(* IEC 61131-3 sources: plcfuzz/testcases/beremiz_projects/random_projects, 27 files *)

(* ---- G4LTL_ST1.st ---- *)
FUNCTION_BLOCK FB_G4LTL

   (* Variable definition *)
   VAR_INPUT
      x0	: BOOL;
      x1	: BOOL;
   END_VAR
   VAR_OUTPUT
      y0	: BOOL;
   END_VAR
   VAR
   (* The total number of states equals to 1 *)
      cstate0	: LINT := 0;
   END_VAR

   (* Control logic *)
CASE cstate0 OF
0:
    IF ((x0 = FALSE) AND  ( TRUE )) OR ((x0 = TRUE) AND  (x1 = TRUE)) THEN
        cstate0 := 0; y0 := FALSE;
    ELSIF ((x0 = TRUE) AND  (x1 = FALSE)) THEN
        cstate0 := 0; y0 := TRUE;
    END_IF;
END_CASE;

END_FUNCTION_BLOCK

(* ---- G4LTL_ST10.st ---- *)
FUNCTION_BLOCK FB_G4LTL

   (* Variable definition *)
   VAR_INPUT
      x1	: BOOL;
      x2	: BOOL;
   END_VAR
   VAR_OUTPUT
      y0	: BOOL;
      y1	: BOOL;
      y2	: BOOL;
   END_VAR
   VAR
   (* The total number of states equals to 6 *)
      cstate79	: LINT := 0;
   END_VAR

   (* Control logic *)
CASE cstate79 OF
0:
    IF ((x1 = FALSE) AND  (x2 = TRUE)) THEN
        cstate79 := 1; y0 := FALSE; y1 := FALSE; y2 := TRUE;
    ELSIF ((x1 = FALSE) AND  (x2 = FALSE)) THEN
        cstate79 := 2; y0 := FALSE; y1 := FALSE; y2 := TRUE;
    ELSIF ((x1 = TRUE) AND  (x2 = FALSE)) THEN
        cstate79 := 3; y0 := TRUE; y1 := TRUE; y2 := FALSE;
    ELSIF ((x1 = TRUE) AND  (x2 = TRUE)) THEN
        cstate79 := 5; y0 := FALSE; y1 := FALSE; y2 := FALSE;
    END_IF;
1:
    IF ((x1 = TRUE) AND  (x2 = FALSE)) THEN
        cstate79 := 3; y0 := TRUE; y1 := TRUE; y2 := FALSE;
    ELSIF ((x1 = TRUE) AND  (x2 = TRUE)) THEN
        cstate79 := 5; y0 := FALSE; y1 := FALSE; y2 := FALSE;
    ELSIF ((x1 = FALSE) AND  ( TRUE )) THEN
        cstate79 := 1; y0 := FALSE; y1 := FALSE; y2 := TRUE;
    END_IF;
2:
    IF ((x1 = TRUE) AND  (x2 = FALSE)) THEN
        cstate79 := 3; y0 := TRUE; y1 := TRUE; y2 := FALSE;
    ELSIF ((x1 = FALSE) AND  (x2 = TRUE)) THEN
        cstate79 := 1; y0 := FALSE; y1 := FALSE; y2 := TRUE;
    ELSIF ((x1 = TRUE) AND  (x2 = TRUE)) THEN
        cstate79 := 5; y0 := FALSE; y1 := FALSE; y2 := FALSE;
    ELSIF ((x1 = FALSE) AND  (x2 = FALSE)) THEN
        cstate79 := 2; y0 := FALSE; y1 := FALSE; y2 := TRUE;
    END_IF;
3:
    IF ((x1 = FALSE) AND  (x2 = TRUE)) THEN
        cstate79 := 4; y0 := FALSE; y1 := FALSE; y2 := TRUE;
    ELSIF (( TRUE ) AND  (x2 = FALSE)) THEN
        cstate79 := 3; y0 := TRUE; y1 := TRUE; y2 := FALSE;
    ELSIF ((x1 = TRUE) AND  (x2 = TRUE)) THEN
        cstate79 := 5; y0 := FALSE; y1 := FALSE; y2 := FALSE;
    END_IF;
4:
    IF ((x1 = TRUE) AND  (x2 = FALSE)) THEN
        cstate79 := 3; y0 := TRUE; y1 := TRUE; y2 := FALSE;
    ELSIF ((x1 = TRUE) AND  (x2 = TRUE)) THEN
        cstate79 := 5; y0 := FALSE; y1 := FALSE; y2 := FALSE;
    ELSIF ((x1 = FALSE) AND  ( TRUE )) THEN
        cstate79 := 4; y0 := FALSE; y1 := FALSE; y2 := TRUE;
    END_IF;
5:
    IF ((x1 = FALSE) AND  (x2 = FALSE)) THEN
        cstate79 := 5; y0 := FALSE; y1 := FALSE; y2 := FALSE;
    ELSIF ((x1 = TRUE) AND  (x2 = TRUE)) THEN
        cstate79 := 5; y0 := FALSE; y1 := FALSE; y2 := FALSE;
    ELSIF ((x1 = TRUE) AND  (x2 = FALSE)) THEN
        cstate79 := 3; y0 := TRUE; y1 := TRUE; y2 := FALSE;
    ELSIF ((x1 = FALSE) AND  (x2 = TRUE)) THEN
        cstate79 := 4; y0 := FALSE; y1 := FALSE; y2 := TRUE;
    END_IF;
END_CASE;

END_FUNCTION_BLOCK

(* ---- G4LTL_ST2.st ---- *)
FUNCTION_BLOCK FB_G4LTL

   (* Variable definition *)
   VAR_INPUT
      x0	: BOOL;
      x1	: BOOL;
   END_VAR
   VAR_OUTPUT
      y0	: BOOL;
   END_VAR
   VAR
   (* The total number of states equals to 1 *)
      cstate99	: LINT := 0;
   END_VAR

   (* Control logic *)
CASE cstate99 OF
0:
    IF ((x0 = FALSE) AND  (x1 = TRUE)) OR ((x0 = TRUE) AND  (x1 = FALSE)) THEN
        cstate99 := 0; y0 := FALSE;
    ELSIF ((x0 = FALSE) AND  (x1 = FALSE)) OR ((x0 = TRUE) AND  (x1 = TRUE)) THEN
        cstate99 := 0; y0 := TRUE;
    END_IF;
END_CASE;

END_FUNCTION_BLOCK

(* ---- G4LTL_ST3.st ---- *)
FUNCTION_BLOCK FB_G4LTL

   (* Variable definition *)
   VAR_INPUT
      x0	: BOOL;
      x1	: BOOL;
      x2	: BOOL;
      x3	: BOOL;
   END_VAR
   VAR_OUTPUT
      y0	: BOOL;
   END_VAR
   VAR
   (* The total number of states equals to 12 *)
      cstate33	: LINT := 0;
   END_VAR

   (* Control logic *)
CASE cstate33 OF
22:
    IF ((x0 = TRUE) AND  (x1 = TRUE) AND  (x2 = TRUE) AND  (x3 = FALSE)) THEN
        cstate33 := 247; y0 := FALSE;
    ELSIF ((x0 = FALSE) AND  ( TRUE ) AND  ( TRUE ) AND  ( TRUE )) OR ((x0 = TRUE) AND  ( TRUE ) AND  (x2 = FALSE) AND  ( TRUE )) THEN
        cstate33 := 22; y0 := FALSE;
    ELSIF ((x0 = TRUE) AND  (x1 = FALSE) AND  (x2 = TRUE) AND  (x3 = FALSE)) THEN
        cstate33 := 246; y0 := TRUE;
    ELSIF ((x0 = TRUE) AND  ( TRUE ) AND  (x2 = TRUE) AND  (x3 = TRUE)) THEN
        cstate33 := 29; y0 := FALSE;
    END_IF;
0:
    IF ((x0 = FALSE) AND  (x1 = FALSE) AND  (x2 = TRUE) AND  (x3 = FALSE)) THEN
        cstate33 := 0; y0 := FALSE;
    ELSIF ((x0 = FALSE) AND  (x1 = TRUE) AND  (x2 = TRUE) AND  (x3 = FALSE)) THEN
        cstate33 := 24; y0 := FALSE;
    ELSIF ((x0 = FALSE) AND  (x1 = TRUE) AND  ( TRUE ) AND  (x3 = TRUE)) OR ((x0 = TRUE) AND  (x1 = TRUE) AND  (x2 = FALSE) AND  (x3 = TRUE)) THEN
        cstate33 := 22; y0 := FALSE;
    ELSIF ((x0 = TRUE) AND  (x1 = TRUE) AND  (x2 = TRUE) AND  (x3 = FALSE)) THEN
        cstate33 := 28; y0 := FALSE;
    ELSIF (( TRUE ) AND  (x1 = TRUE) AND  (x2 = FALSE) AND  (x3 = FALSE)) THEN
        cstate33 := 20; y0 := FALSE;
    ELSIF ((x0 = TRUE) AND  (x1 = FALSE) AND  (x2 = TRUE) AND  (x3 = FALSE)) THEN
        cstate33 := 27; y0 := TRUE;
    ELSIF ((x0 = TRUE) AND  (x1 = TRUE) AND  (x2 = TRUE) AND  (x3 = TRUE)) THEN
        cstate33 := 29; y0 := FALSE;
    ELSIF (( TRUE ) AND  (x1 = FALSE) AND  (x2 = FALSE) AND  ( TRUE )) OR (( TRUE ) AND  (x1 = FALSE) AND  (x2 = TRUE) AND  (x3 = TRUE)) THEN
        cstate33 := 18; y0 := FALSE;
    END_IF;
243:
    IF ((x0 = FALSE) AND  (x1 = FALSE) AND  (x2 = TRUE) AND  (x3 = TRUE)) OR ((x0 = TRUE) AND  ( TRUE ) AND  (x2 = TRUE) AND  (x3 = TRUE)) THEN
        cstate33 := 29; y0 := FALSE;
    ELSIF (( TRUE ) AND  ( TRUE ) AND  (x2 = FALSE) AND  (x3 = FALSE)) THEN
        cstate33 := 20; y0 := FALSE;
    ELSIF ((x0 = FALSE) AND  (x1 = FALSE) AND  (x2 = FALSE) AND  (x3 = TRUE)) OR ((x0 = FALSE) AND  (x1 = TRUE) AND  ( TRUE ) AND  (x3 = TRUE)) OR ((x0 = TRUE) AND  ( TRUE ) AND  (x2 = FALSE) AND  (x3 = TRUE)) THEN
        cstate33 := 22; y0 := FALSE;
    ELSIF ((x0 = FALSE) AND  (x1 = TRUE) AND  (x2 = TRUE) AND  (x3 = FALSE)) THEN
        cstate33 := 24; y0 := FALSE;
    ELSIF ((x0 = TRUE) AND  (x1 = TRUE) AND  (x2 = TRUE) AND  (x3 = FALSE)) THEN
        cstate33 := 28; y0 := FALSE;
    ELSIF (( TRUE ) AND  (x1 = FALSE) AND  (x2 = TRUE) AND  (x3 = FALSE)) THEN
        cstate33 := 243; y0 := TRUE;
    END_IF;
24:
    IF ((x0 = TRUE) AND  ( TRUE ) AND  (x2 = TRUE) AND  (x3 = TRUE)) THEN
        cstate33 := 29; y0 := FALSE;
    ELSIF (( TRUE ) AND  ( TRUE ) AND  (x2 = FALSE) AND  (x3 = FALSE)) THEN
        cstate33 := 20; y0 := FALSE;
    ELSIF ((x0 = FALSE) AND  ( TRUE ) AND  ( TRUE ) AND  (x3 = TRUE)) OR ((x0 = TRUE) AND  ( TRUE ) AND  (x2 = FALSE) AND  (x3 = TRUE)) THEN
        cstate33 := 22; y0 := FALSE;
    ELSIF ((x0 = TRUE) AND  (x1 = TRUE) AND  (x2 = TRUE) AND  (x3 = FALSE)) THEN
        cstate33 := 28; y0 := FALSE;
    ELSIF ((x0 = TRUE) AND  (x1 = FALSE) AND  (x2 = TRUE) AND  (x3 = FALSE)) THEN
        cstate33 := 243; y0 := TRUE;
    ELSIF ((x0 = FALSE) AND  ( TRUE ) AND  (x2 = TRUE) AND  (x3 = FALSE)) THEN
        cstate33 := 24; y0 := FALSE;
    END_IF;
246:
    IF ((x0 = FALSE) AND  (x1 = FALSE) AND  (x2 = FALSE) AND  ( TRUE )) OR ((x0 = FALSE) AND  (x1 = TRUE) AND  (x2 = FALSE) AND  ( TRUE )) OR ((x0 = FALSE) AND  (x1 = TRUE) AND  (x2 = TRUE) AND  (x3 = TRUE)) OR ((x0 = TRUE) AND  ( TRUE ) AND  (x2 = FALSE) AND  ( TRUE )) THEN
        cstate33 := 22; y0 := FALSE;
    ELSIF (( TRUE ) AND  (x1 = FALSE) AND  (x2 = TRUE) AND  (x3 = FALSE)) THEN
        cstate33 := 246; y0 := TRUE;
    ELSIF ((x0 = FALSE) AND  (x1 = FALSE) AND  (x2 = TRUE) AND  (x3 = TRUE)) OR ((x0 = TRUE) AND  ( TRUE ) AND  (x2 = TRUE) AND  (x3 = TRUE)) THEN
        cstate33 := 29; y0 := FALSE;
    ELSIF ((x0 = FALSE) AND  (x1 = TRUE) AND  (x2 = TRUE) AND  (x3 = FALSE)) THEN
        cstate33 := 786; y0 := FALSE;
    ELSIF ((x0 = TRUE) AND  (x1 = TRUE) AND  (x2 = TRUE) AND  (x3 = FALSE)) THEN
        cstate33 := 247; y0 := FALSE;
    END_IF;
27:
    IF ((x0 = FALSE) AND  (x1 = TRUE) AND  (x2 = TRUE) AND  (x3 = FALSE)) THEN
        cstate33 := 24; y0 := FALSE;
    ELSIF (( TRUE ) AND  (x1 = TRUE) AND  (x2 = FALSE) AND  (x3 = FALSE)) THEN
        cstate33 := 20; y0 := FALSE;
    ELSIF ((x0 = FALSE) AND  (x1 = TRUE) AND  ( TRUE ) AND  (x3 = TRUE)) OR ((x0 = TRUE) AND  (x1 = TRUE) AND  (x2 = FALSE) AND  (x3 = TRUE)) THEN
        cstate33 := 22; y0 := FALSE;
    ELSIF ((x0 = TRUE) AND  (x1 = TRUE) AND  (x2 = TRUE) AND  (x3 = FALSE)) THEN
        cstate33 := 28; y0 := FALSE;
    ELSIF (( TRUE ) AND  (x1 = FALSE) AND  (x2 = TRUE) AND  (x3 = FALSE)) THEN
        cstate33 := 27; y0 := TRUE;
    ELSIF ((x0 = TRUE) AND  (x1 = TRUE) AND  (x2 = TRUE) AND  (x3 = TRUE)) THEN
        cstate33 := 29; y0 := FALSE;
    ELSIF (( TRUE ) AND  (x1 = FALSE) AND  (x2 = FALSE) AND  ( TRUE )) OR (( TRUE ) AND  (x1 = FALSE) AND  (x2 = TRUE) AND  (x3 = TRUE)) THEN
        cstate33 := 18; y0 := FALSE;
    END_IF;
247:
    IF ((x0 = FALSE) AND  (x1 = TRUE) AND  (x2 = TRUE) AND  (x3 = FALSE)) THEN
        cstate33 := 786; y0 := FALSE;
    ELSIF ((x0 = FALSE) AND  (x1 = FALSE) AND  (x2 = TRUE) AND  (x3 = FALSE)) OR ((x0 = TRUE) AND  (x1 = TRUE) AND  (x2 = TRUE) AND  (x3 = FALSE)) THEN
        cstate33 := 247; y0 := FALSE;
    ELSIF ((x0 = FALSE) AND  (x1 = FALSE) AND  (x2 = FALSE) AND  ( TRUE )) OR ((x0 = FALSE) AND  (x1 = TRUE) AND  (x2 = FALSE) AND  ( TRUE )) OR ((x0 = FALSE) AND  (x1 = TRUE) AND  (x2 = TRUE) AND  (x3 = TRUE)) OR ((x0 = TRUE) AND  ( TRUE ) AND  (x2 = FALSE) AND  ( TRUE )) THEN
        cstate33 := 22; y0 := FALSE;
    ELSIF ((x0 = TRUE) AND  (x1 = FALSE) AND  (x2 = TRUE) AND  (x3 = FALSE)) THEN
        cstate33 := 246; y0 := TRUE;
    ELSIF ((x0 = FALSE) AND  (x1 = FALSE) AND  (x2 = TRUE) AND  (x3 = TRUE)) OR ((x0 = TRUE) AND  ( TRUE ) AND  (x2 = TRUE) AND  (x3 = TRUE)) THEN
        cstate33 := 29; y0 := FALSE;
    END_IF;
786:
    IF ((x0 = TRUE) AND  (x1 = TRUE) AND  (x2 = TRUE) AND  (x3 = FALSE)) THEN
        cstate33 := 247; y0 := FALSE;
    ELSIF ((x0 = FALSE) AND  ( TRUE ) AND  (x2 = FALSE) AND  ( TRUE )) OR ((x0 = FALSE) AND  ( TRUE ) AND  (x2 = TRUE) AND  (x3 = TRUE)) OR ((x0 = TRUE) AND  ( TRUE ) AND  (x2 = FALSE) AND  ( TRUE )) THEN
        cstate33 := 22; y0 := FALSE;
    ELSIF ((x0 = FALSE) AND  ( TRUE ) AND  (x2 = TRUE) AND  (x3 = FALSE)) THEN
        cstate33 := 786; y0 := FALSE;
    ELSIF ((x0 = TRUE) AND  (x1 = FALSE) AND  (x2 = TRUE) AND  (x3 = FALSE)) THEN
        cstate33 := 246; y0 := TRUE;
    ELSIF ((x0 = TRUE) AND  ( TRUE ) AND  (x2 = TRUE) AND  (x3 = TRUE)) THEN
        cstate33 := 29; y0 := FALSE;
    END_IF;
28:
    IF ((x0 = FALSE) AND  (x1 = FALSE) AND  (x2 = TRUE) AND  (x3 = FALSE)) OR ((x0 = TRUE) AND  (x1 = TRUE) AND  (x2 = TRUE) AND  (x3 = FALSE)) THEN
        cstate33 := 28; y0 := FALSE;
    ELSIF (( TRUE ) AND  ( TRUE ) AND  (x2 = FALSE) AND  (x3 = FALSE)) THEN
        cstate33 := 20; y0 := FALSE;
    ELSIF ((x0 = FALSE) AND  (x1 = FALSE) AND  (x2 = FALSE) AND  (x3 = TRUE)) OR ((x0 = FALSE) AND  (x1 = TRUE) AND  ( TRUE ) AND  (x3 = TRUE)) OR ((x0 = TRUE) AND  ( TRUE ) AND  (x2 = FALSE) AND  (x3 = TRUE)) THEN
        cstate33 := 22; y0 := FALSE;
    ELSIF ((x0 = FALSE) AND  (x1 = TRUE) AND  (x2 = TRUE) AND  (x3 = FALSE)) THEN
        cstate33 := 24; y0 := FALSE;
    ELSIF ((x0 = TRUE) AND  (x1 = FALSE) AND  (x2 = TRUE) AND  (x3 = FALSE)) THEN
        cstate33 := 243; y0 := TRUE;
    ELSIF ((x0 = FALSE) AND  (x1 = FALSE) AND  (x2 = TRUE) AND  (x3 = TRUE)) OR ((x0 = TRUE) AND  ( TRUE ) AND  (x2 = TRUE) AND  (x3 = TRUE)) THEN
        cstate33 := 29; y0 := FALSE;
    END_IF;
29:
    IF ((x0 = TRUE) AND  (x1 = TRUE) AND  (x2 = TRUE) AND  (x3 = FALSE)) THEN
        cstate33 := 247; y0 := FALSE;
    ELSIF ((x0 = FALSE) AND  (x1 = FALSE) AND  (x2 = TRUE) AND  ( TRUE )) OR ((x0 = TRUE) AND  ( TRUE ) AND  (x2 = TRUE) AND  (x3 = TRUE)) THEN
        cstate33 := 29; y0 := FALSE;
    ELSIF ((x0 = TRUE) AND  (x1 = FALSE) AND  (x2 = TRUE) AND  (x3 = FALSE)) THEN
        cstate33 := 246; y0 := TRUE;
    ELSIF ((x0 = FALSE) AND  (x1 = FALSE) AND  (x2 = FALSE) AND  ( TRUE )) OR ((x0 = FALSE) AND  (x1 = TRUE) AND  ( TRUE ) AND  ( TRUE )) OR ((x0 = TRUE) AND  ( TRUE ) AND  (x2 = FALSE) AND  ( TRUE )) THEN
        cstate33 := 22; y0 := FALSE;
    END_IF;
18:
    IF ((x0 = TRUE) AND  (x1 = TRUE) AND  (x2 = TRUE) AND  (x3 = TRUE)) THEN
        cstate33 := 29; y0 := FALSE;
    ELSIF ((x0 = TRUE) AND  (x1 = FALSE) AND  (x2 = TRUE) AND  (x3 = FALSE)) THEN
        cstate33 := 27; y0 := TRUE;
    ELSIF ((x0 = FALSE) AND  (x1 = FALSE) AND  ( TRUE ) AND  ( TRUE )) OR ((x0 = TRUE) AND  (x1 = FALSE) AND  (x2 = FALSE) AND  ( TRUE )) OR ((x0 = TRUE) AND  (x1 = FALSE) AND  (x2 = TRUE) AND  (x3 = TRUE)) THEN
        cstate33 := 18; y0 := FALSE;
    ELSIF ((x0 = FALSE) AND  (x1 = TRUE) AND  ( TRUE ) AND  (x3 = FALSE)) OR ((x0 = TRUE) AND  (x1 = TRUE) AND  (x2 = FALSE) AND  (x3 = FALSE)) THEN
        cstate33 := 20; y0 := FALSE;
    ELSIF ((x0 = FALSE) AND  (x1 = TRUE) AND  ( TRUE ) AND  (x3 = TRUE)) OR ((x0 = TRUE) AND  (x1 = TRUE) AND  (x2 = FALSE) AND  (x3 = TRUE)) THEN
        cstate33 := 22; y0 := FALSE;
    ELSIF ((x0 = TRUE) AND  (x1 = TRUE) AND  (x2 = TRUE) AND  (x3 = FALSE)) THEN
        cstate33 := 28; y0 := FALSE;
    END_IF;
20:
    IF ((x0 = TRUE) AND  ( TRUE ) AND  (x2 = TRUE) AND  (x3 = TRUE)) THEN
        cstate33 := 29; y0 := FALSE;
    ELSIF ((x0 = FALSE) AND  ( TRUE ) AND  ( TRUE ) AND  (x3 = TRUE)) OR ((x0 = TRUE) AND  ( TRUE ) AND  (x2 = FALSE) AND  (x3 = TRUE)) THEN
        cstate33 := 22; y0 := FALSE;
    ELSIF ((x0 = FALSE) AND  ( TRUE ) AND  ( TRUE ) AND  (x3 = FALSE)) OR ((x0 = TRUE) AND  ( TRUE ) AND  (x2 = FALSE) AND  (x3 = FALSE)) THEN
        cstate33 := 20; y0 := FALSE;
    ELSIF ((x0 = TRUE) AND  (x1 = TRUE) AND  (x2 = TRUE) AND  (x3 = FALSE)) THEN
        cstate33 := 28; y0 := FALSE;
    ELSIF ((x0 = TRUE) AND  (x1 = FALSE) AND  (x2 = TRUE) AND  (x3 = FALSE)) THEN
        cstate33 := 243; y0 := TRUE;
    END_IF;
END_CASE;

END_FUNCTION_BLOCK

(* ---- G4LTL_ST4.st ---- *)
FUNCTION_BLOCK FB_G4LTL

   (* Variable definition *)
   VAR_INPUT
      x0	: BOOL;
      x1	: BOOL;
      x2	: BOOL;
      x3	: BOOL;
   END_VAR
   VAR_OUTPUT
      y0	: BOOL;
      y1	: BOOL;
   END_VAR
   VAR
   (* The total number of states equals to 2 *)
      cstate29	: LINT := 0;
   END_VAR

   (* Control logic *)
CASE cstate29 OF
0:
    IF ((x0 = FALSE) AND  (x1 = FALSE) AND  (x2 = FALSE) AND  (x3 = TRUE)) THEN
        cstate29 := 0; y0 := FALSE; y1 := FALSE;
    ELSIF ((x0 = FALSE) AND  (x1 = TRUE) AND  ( TRUE ) AND  (x3 = TRUE)) OR ((x0 = TRUE) AND  (x1 = FALSE) AND  (x2 = TRUE) AND  ( TRUE )) OR ((x0 = TRUE) AND  (x1 = TRUE) AND  (x2 = FALSE) AND  (x3 = TRUE)) OR ((x0 = TRUE) AND  (x1 = TRUE) AND  (x2 = TRUE) AND  ( TRUE )) THEN
        cstate29 := 1; y0 := FALSE; y1 := FALSE;
    ELSIF ((x0 = FALSE) AND  (x1 = FALSE) AND  (x2 = FALSE) AND  (x3 = FALSE)) OR ((x0 = FALSE) AND  (x1 = FALSE) AND  (x2 = TRUE) AND  ( TRUE )) OR ((x0 = FALSE) AND  (x1 = TRUE) AND  ( TRUE ) AND  (x3 = FALSE)) THEN
        cstate29 := 0; y0 := FALSE; y1 := FALSE;
    ELSIF ((x0 = TRUE) AND  (x1 = TRUE) AND  (x2 = FALSE) AND  (x3 = FALSE)) THEN
        cstate29 := 0; y0 := TRUE; y1 := TRUE;
    ELSIF ((x0 = TRUE) AND  (x1 = FALSE) AND  (x2 = FALSE) AND  (x3 = TRUE)) THEN
        cstate29 := 0; y0 := TRUE; y1 := FALSE;
    ELSIF ((x0 = TRUE) AND  (x1 = FALSE) AND  (x2 = FALSE) AND  (x3 = FALSE)) THEN
        cstate29 := 0; y0 := TRUE; y1 := FALSE;
    END_IF;
1:
    IF ((x0 = TRUE) AND  (x1 = FALSE) AND  (x2 = FALSE) AND  ( TRUE )) OR ((x0 = TRUE) AND  (x1 = TRUE) AND  (x2 = FALSE) AND  (x3 = FALSE)) THEN
        cstate29 := 1; y0 := FALSE; y1 := FALSE;
    ELSIF ((x0 = FALSE) AND  (x1 = FALSE) AND  (x2 = FALSE) AND  (x3 = FALSE)) OR ((x0 = FALSE) AND  (x1 = FALSE) AND  (x2 = TRUE) AND  ( TRUE )) OR ((x0 = FALSE) AND  (x1 = TRUE) AND  ( TRUE ) AND  (x3 = FALSE)) THEN
        cstate29 := 1; y0 := FALSE; y1 := FALSE;
    ELSIF ((x0 = FALSE) AND  (x1 = TRUE) AND  ( TRUE ) AND  (x3 = TRUE)) OR ((x0 = TRUE) AND  (x1 = FALSE) AND  (x2 = TRUE) AND  ( TRUE )) OR ((x0 = TRUE) AND  (x1 = TRUE) AND  (x2 = FALSE) AND  (x3 = TRUE)) OR ((x0 = TRUE) AND  (x1 = TRUE) AND  (x2 = TRUE) AND  ( TRUE )) THEN
        cstate29 := 1; y0 := FALSE; y1 := FALSE;
    ELSIF ((x0 = FALSE) AND  (x1 = FALSE) AND  (x2 = FALSE) AND  (x3 = TRUE)) THEN
        cstate29 := 1; y0 := FALSE; y1 := FALSE;
    END_IF;
END_CASE;

END_FUNCTION_BLOCK

(* ---- G4LTL_ST5.st ---- *)
FUNCTION_BLOCK FB_G4LTL

   (* Variable definition *)
   VAR_INPUT
      x0	: BOOL;
      x1	: BOOL;
      c1_geq500	: BOOL;
   END_VAR
   VAR_OUTPUT
      y0	: BOOL;
      c1_add1	: BOOL;
      c1_reset	: BOOL;
   END_VAR
   VAR
   (* The total number of states equals to 4 *)
      cstate69	: LINT := 0;
   END_VAR

   (* Control logic *)
CASE cstate69 OF
0:
    IF ((x0 = FALSE) AND  (x1 = TRUE) AND  (c1_geq500 = TRUE)) THEN
        cstate69 := 3; y0 := TRUE; c1_add1 := FALSE; c1_reset := TRUE;
    ELSIF ((x0 = FALSE) AND  (x1 = FALSE) AND  (c1_geq500 = TRUE)) THEN
        cstate69 := 3; y0 := TRUE; c1_add1 := FALSE; c1_reset := FALSE;
    ELSIF ((x0 = FALSE) AND  (x1 = TRUE) AND  (c1_geq500 = FALSE)) THEN
        cstate69 := 3; y0 := FALSE; c1_add1 := FALSE; c1_reset := TRUE;
    ELSIF ((x0 = FALSE) AND  (x1 = FALSE) AND  (c1_geq500 = FALSE)) THEN
        cstate69 := 3; y0 := FALSE; c1_add1 := FALSE; c1_reset := FALSE;
    ELSIF ((x0 = TRUE) AND  (x1 = TRUE) AND  ( TRUE )) THEN
        cstate69 := 1; y0 := FALSE; c1_add1 := FALSE; c1_reset := FALSE;
    ELSIF ((x0 = TRUE) AND  (x1 = FALSE) AND  (c1_geq500 = TRUE)) THEN
        cstate69 := 2; y0 := TRUE; c1_add1 := TRUE; c1_reset := FALSE;
    ELSIF ((x0 = TRUE) AND  (x1 = FALSE) AND  (c1_geq500 = FALSE)) THEN
        cstate69 := 2; y0 := FALSE; c1_add1 := TRUE; c1_reset := FALSE;
    END_IF;
1:
    IF ((x0 = TRUE) AND  (x1 = TRUE) AND  ( TRUE )) THEN
        cstate69 := 1; y0 := FALSE; c1_add1 := FALSE; c1_reset := FALSE;
    ELSIF ((x0 = FALSE) AND  ( TRUE ) AND  (c1_geq500 = FALSE)) OR ((x0 = TRUE) AND  (x1 = FALSE) AND  (c1_geq500 = FALSE)) THEN
        cstate69 := 1; y0 := FALSE; c1_add1 := FALSE; c1_reset := FALSE;
    ELSIF ((x0 = FALSE) AND  ( TRUE ) AND  (c1_geq500 = TRUE)) OR ((x0 = TRUE) AND  (x1 = FALSE) AND  (c1_geq500 = TRUE)) THEN
        cstate69 := 1; y0 := FALSE; c1_add1 := FALSE; c1_reset := FALSE;
    END_IF;
2:
    IF ((x0 = TRUE) AND  (x1 = TRUE) AND  ( TRUE )) THEN
        cstate69 := 1; y0 := FALSE; c1_add1 := FALSE; c1_reset := FALSE;
    ELSIF ((x0 = FALSE) AND  (x1 = FALSE) AND  (c1_geq500 = TRUE)) THEN
        cstate69 := 3; y0 := TRUE; c1_add1 := FALSE; c1_reset := FALSE;
    ELSIF ((x0 = FALSE) AND  (x1 = TRUE) AND  (c1_geq500 = FALSE)) THEN
        cstate69 := 3; y0 := FALSE; c1_add1 := FALSE; c1_reset := TRUE;
    ELSIF ((x0 = FALSE) AND  (x1 = TRUE) AND  (c1_geq500 = TRUE)) THEN
        cstate69 := 3; y0 := TRUE; c1_add1 := FALSE; c1_reset := TRUE;
    ELSIF ((x0 = FALSE) AND  (x1 = FALSE) AND  (c1_geq500 = FALSE)) THEN
        cstate69 := 3; y0 := FALSE; c1_add1 := FALSE; c1_reset := FALSE;
    ELSIF ((x0 = TRUE) AND  (x1 = FALSE) AND  (c1_geq500 = FALSE)) THEN
        cstate69 := 2; y0 := FALSE; c1_add1 := FALSE; c1_reset := FALSE;
    ELSIF ((x0 = TRUE) AND  (x1 = FALSE) AND  (c1_geq500 = TRUE)) THEN
        cstate69 := 2; y0 := TRUE; c1_add1 := FALSE; c1_reset := FALSE;
    END_IF;
3:
    IF ((x0 = FALSE) AND  (x1 = FALSE) AND  (c1_geq500 = FALSE)) THEN
        cstate69 := 3; y0 := FALSE; c1_add1 := FALSE; c1_reset := FALSE;
    ELSIF ((x0 = FALSE) AND  (x1 = FALSE) AND  (c1_geq500 = TRUE)) THEN
        cstate69 := 3; y0 := TRUE; c1_add1 := FALSE; c1_reset := FALSE;
    ELSIF ((x0 = FALSE) AND  (x1 = TRUE) AND  (c1_geq500 = FALSE)) THEN
        cstate69 := 3; y0 := FALSE; c1_add1 := FALSE; c1_reset := TRUE;
    ELSIF ((x0 = FALSE) AND  (x1 = TRUE) AND  (c1_geq500 = TRUE)) THEN
        cstate69 := 3; y0 := TRUE; c1_add1 := FALSE; c1_reset := TRUE;
    ELSIF ((x0 = TRUE) AND  (x1 = TRUE) AND  ( TRUE )) THEN
        cstate69 := 1; y0 := FALSE; c1_add1 := FALSE; c1_reset := FALSE;
    ELSIF ((x0 = TRUE) AND  (x1 = FALSE) AND  (c1_geq500 = FALSE)) THEN
        cstate69 := 2; y0 := FALSE; c1_add1 := TRUE; c1_reset := FALSE;
    ELSIF ((x0 = TRUE) AND  (x1 = FALSE) AND  (c1_geq500 = TRUE)) THEN
        cstate69 := 2; y0 := TRUE; c1_add1 := TRUE; c1_reset := FALSE;
    END_IF;
END_CASE;

END_FUNCTION_BLOCK

(* ---- G4LTL_ST6.st ---- *)
FUNCTION_BLOCK FB_G4LTL

   (* Variable definition *)
   VAR_INPUT
      x1	: BOOL;
   END_VAR
   VAR_OUTPUT
      y1	: BOOL;
   END_VAR
   VAR
   (* The total number of states equals to 7 *)
      cstate14	: LINT := 0;
      t	: TON;
      t_reset	: BOOL := FALSE;
      t_up	: BOOL := FALSE;
      t_start	: BOOL := FALSE;
   END_VAR

   (* Constant definition (depending on compiler, one might need to move to normal variables) *)

   (* Each time constant has a difference of 1 period (cycle-time); please substract it when needed  *)
   VAR CONST
      T_VALUE	: TIME := TIME#5s;
   END_VAR

   (* Control logic *)
CASE cstate14 OF
0:
    IF ((x1 = FALSE) AND  (t.Q = FALSE)) THEN
        cstate14 := 1; y1 := FALSE; t_start := FALSE;
    ELSIF ((x1 = TRUE) AND  ( TRUE )) THEN
        cstate14 := 3; y1 := TRUE; t_start := FALSE;
    ELSIF ((x1 = FALSE) AND  (t.Q = TRUE)) THEN
        cstate14 := 5; y1 := FALSE; t_start := FALSE;
    END_IF;
1:
    IF ((x1 = FALSE) AND  (t.Q = FALSE)) THEN
        cstate14 := 1; y1 := FALSE; t_start := FALSE;
    ELSIF ((x1 = FALSE) AND  (t.Q = TRUE)) THEN
        cstate14 := 5; y1 := FALSE; t_start := FALSE;
    ELSIF ((x1 = TRUE) AND  ( TRUE )) THEN
        cstate14 := 3; y1 := TRUE; t_start := FALSE;
    END_IF;
2:
    IF ((x1 = TRUE) AND  (t.Q = FALSE)) THEN
        cstate14 := 2; y1 := TRUE; t_start := FALSE;
    ELSIF ((x1 = TRUE) AND  (t.Q = TRUE)) THEN
        cstate14 := 3; y1 := TRUE; t_start := FALSE;
    ELSIF ((x1 = FALSE) AND  (t.Q = FALSE)) THEN
        cstate14 := 4; y1 := TRUE; t_start := TRUE; t_up := FALSE;
    ELSIF ((x1 = FALSE) AND  (t.Q = TRUE)) THEN
        cstate14 := 6; y1 := TRUE; t_start := TRUE; t_up := FALSE;
    END_IF;
3:
    IF ((x1 = FALSE) AND  (t.Q = TRUE)) THEN
        cstate14 := 6; y1 := TRUE; t_start := TRUE; t_up := FALSE;
    ELSIF ((x1 = FALSE) AND  (t.Q = FALSE)) THEN
        cstate14 := 4; y1 := TRUE; t_start := TRUE; t_up := FALSE;
    ELSIF ((x1 = TRUE) AND  ( TRUE )) THEN
        cstate14 := 3; y1 := TRUE; t_start := FALSE;
    END_IF;
4:
    IF ((x1 = FALSE) AND  (t.Q = TRUE)) THEN
        cstate14 := 5; y1 := FALSE; t_start := FALSE;
    ELSIF ((x1 = FALSE) AND  (t.Q = FALSE)) THEN
        cstate14 := 4; y1 := TRUE; t_start := FALSE;
    ELSIF ((x1 = TRUE) AND  (t.Q = FALSE)) THEN
        cstate14 := 2; y1 := TRUE; t_start := FALSE;
    ELSIF ((x1 = TRUE) AND  (t.Q = TRUE)) THEN
        cstate14 := 3; y1 := TRUE; t_start := FALSE;
    END_IF;
5:
    IF ((x1 = TRUE) AND  ( TRUE )) THEN
        cstate14 := 3; y1 := TRUE; t_start := FALSE;
    ELSIF ((x1 = FALSE) AND  (t.Q = FALSE)) THEN
        cstate14 := 1; y1 := FALSE; t_start := FALSE;
    ELSIF ((x1 = FALSE) AND  (t.Q = TRUE)) THEN
        cstate14 := 5; y1 := FALSE; t_start := FALSE;
    END_IF;
6:
    IF ((x1 = FALSE) AND  (t.Q = TRUE)) THEN
        cstate14 := 5; y1 := FALSE; t_start := FALSE;
    ELSIF ((x1 = FALSE) AND  (t.Q = FALSE)) THEN
        cstate14 := 4; y1 := TRUE; t_start := FALSE;
    ELSIF ((x1 = TRUE) AND  (t.Q = FALSE)) THEN
        cstate14 := 2; y1 := TRUE; t_start := FALSE;
    ELSIF ((x1 = TRUE) AND  (t.Q = TRUE)) THEN
        cstate14 := 3; y1 := TRUE; t_start := FALSE;
    END_IF;
END_CASE;

(* Additional processing to handle clocks - in CODESYS, it only starts
    with rising edge and can not be placed inside IF statement *)
IF(t_up = TRUE) THEN
    t_reset := TRUE;
ELSIF(t_start = TRUE AND t_up = FALSE) THEN
    t_up := TRUE;  t_reset := FALSE;
END_IF
t(IN:=t_reset, PT:=T_VALUE);

END_FUNCTION_BLOCK

(* ---- G4LTL_ST7.st ---- *)
FUNCTION_BLOCK FB_G4LTL

   (* Variable definition *)
   VAR_INPUT
      x1	: BOOL;
   END_VAR
   VAR_OUTPUT
      y1	: BOOL;
   END_VAR
   VAR
   (* The total number of states equals to 7 *)
      cstate58	: LINT := 0;
      t	: TON;
      t_reset	: BOOL := FALSE;
      t_up	: BOOL := FALSE;
      t_start	: BOOL := FALSE;
   END_VAR

   (* Constant definition (depending on compiler, one might need to move to normal variables) *)

   (* Each time constant has a difference of 1 period (cycle-time); please substract it when needed  *)
   VAR CONST
      T_VALUE	: TIME := TIME#3s;
   END_VAR

   (* Control logic *)
CASE cstate58 OF
0:
    IF ((x1 = TRUE) AND  (t.Q = FALSE)) THEN
        cstate58 := 2; y1 := FALSE; t_start := FALSE;
    ELSIF ((x1 = FALSE) AND  ( TRUE )) THEN
        cstate58 := 6; y1 := FALSE; t_start := FALSE;
    ELSIF ((x1 = TRUE) AND  (t.Q = TRUE)) THEN
        cstate58 := 2; y1 := TRUE; t_start := FALSE;
    END_IF;
1:
    IF ((x1 = TRUE) AND  (t.Q = TRUE)) THEN
        cstate58 := 2; y1 := TRUE; t_start := FALSE;
    ELSIF ((x1 = TRUE) AND  (t.Q = FALSE)) THEN
        cstate58 := 1; y1 := FALSE; t_start := FALSE;
    ELSIF ((x1 = FALSE) AND  (t.Q = TRUE)) THEN
        cstate58 := 6; y1 := FALSE; t_start := FALSE;
    ELSIF ((x1 = FALSE) AND  (t.Q = FALSE)) THEN
        cstate58 := 5; y1 := FALSE; t_start := FALSE;
    END_IF;
2:
    IF ((x1 = TRUE) AND  (t.Q = FALSE)) THEN
        cstate58 := 2; y1 := FALSE; t_start := FALSE;
    ELSIF ((x1 = TRUE) AND  (t.Q = TRUE)) THEN
        cstate58 := 2; y1 := TRUE; t_start := FALSE;
    ELSIF ((x1 = FALSE) AND  ( TRUE )) THEN
        cstate58 := 6; y1 := FALSE; t_start := FALSE;
    END_IF;
3:
    IF ((x1 = TRUE) AND  (t.Q = FALSE)) THEN
        cstate58 := 3; y1 := FALSE; t_start := FALSE;
    ELSIF ((x1 = FALSE) AND  (t.Q = FALSE)) THEN
        cstate58 := 4; y1 := FALSE; t_start := FALSE;
    ELSIF ((x1 = TRUE) AND  (t.Q = TRUE)) THEN
        cstate58 := 2; y1 := TRUE; t_start := FALSE;
    ELSIF ((x1 = FALSE) AND  (t.Q = TRUE)) THEN
        cstate58 := 6; y1 := FALSE; t_start := FALSE;
    END_IF;
4:
    IF ((x1 = FALSE) AND  (t.Q = FALSE)) THEN
        cstate58 := 4; y1 := FALSE; t_start := FALSE;
    ELSIF ((x1 = FALSE) AND  (t.Q = TRUE)) THEN
        cstate58 := 6; y1 := FALSE; t_start := FALSE;
    ELSIF ((x1 = TRUE) AND  (t.Q = FALSE)) THEN
        cstate58 := 3; y1 := FALSE; t_start := TRUE; t_up := FALSE;
    ELSIF ((x1 = TRUE) AND  (t.Q = TRUE)) THEN
        cstate58 := 1; y1 := TRUE; t_start := TRUE; t_up := FALSE;
    END_IF;
5:
    IF ((x1 = FALSE) AND  (t.Q = TRUE)) THEN
        cstate58 := 6; y1 := FALSE; t_start := FALSE;
    ELSIF ((x1 = FALSE) AND  (t.Q = FALSE)) THEN
        cstate58 := 5; y1 := FALSE; t_start := FALSE;
    ELSIF ((x1 = TRUE) AND  (t.Q = TRUE)) THEN
        cstate58 := 1; y1 := TRUE; t_start := TRUE; t_up := FALSE;
    ELSIF ((x1 = TRUE) AND  (t.Q = FALSE)) THEN
        cstate58 := 3; y1 := FALSE; t_start := TRUE; t_up := FALSE;
    END_IF;
6:
    IF ((x1 = TRUE) AND  (t.Q = TRUE)) THEN
        cstate58 := 1; y1 := TRUE; t_start := TRUE; t_up := FALSE;
    ELSIF ((x1 = TRUE) AND  (t.Q = FALSE)) THEN
        cstate58 := 3; y1 := FALSE; t_start := TRUE; t_up := FALSE;
    ELSIF ((x1 = FALSE) AND  ( TRUE )) THEN
        cstate58 := 6; y1 := FALSE; t_start := FALSE;
    END_IF;
END_CASE;

(* Additional processing to handle clocks - in CODESYS, it only starts
    with rising edge and can not be placed inside IF statement *)
IF(t_up = TRUE) THEN
    t_reset := TRUE;
ELSIF(t_start = TRUE AND t_up = FALSE) THEN
    t_up := TRUE;  t_reset := FALSE;
END_IF
t(IN:=t_reset, PT:=T_VALUE);

END_FUNCTION_BLOCK

(* ---- G4LTL_ST8.st ---- *)
FUNCTION_BLOCK FB_G4LTL

   (* Variable definition *)
   VAR_INPUT
      x1	: BOOL;
   END_VAR
   VAR_OUTPUT
      y1	: BOOL;
   END_VAR
   VAR
   (* The total number of states equals to 18 *)
      cstate83	: LINT := 0;
      t0	: TON;
      t0_reset	: BOOL := FALSE;
      t0_up	: BOOL := FALSE;
      t0_start	: BOOL := FALSE;
      t1	: TON;
      t1_reset	: BOOL := FALSE;
      t1_up	: BOOL := FALSE;
      t1_start	: BOOL := FALSE;
   END_VAR

   (* Constant definition (depending on compiler, one might need to move to normal variables) *)

   (* Each time constant has a difference of 1 period (cycle-time); please substract it when needed  *)
   VAR CONST
      T0_VALUE	: TIME := TIME#5s;
      T1_VALUE	: TIME := TIME#3s;
   END_VAR

   (* Control logic *)
CASE cstate83 OF
11:
    IF ((x1 = FALSE) AND  (t0.Q = TRUE) AND  (t1.Q = TRUE)) THEN
        cstate83 := 14; y1 := TRUE; t0_start := FALSE;t1_start := TRUE; t1_up := FALSE;
    ELSIF ((x1 = TRUE) AND  (t0.Q = TRUE) AND  ( TRUE )) THEN
        cstate83 := 10; y1 := FALSE; t0_start := FALSE;t1_start := FALSE;
    ELSIF ((x1 = TRUE) AND  (t0.Q = FALSE) AND  ( TRUE )) THEN
        cstate83 := 11; y1 := FALSE; t0_start := FALSE;t1_start := FALSE;
    ELSIF ((x1 = FALSE) AND  (t0.Q = TRUE) AND  (t1.Q = FALSE)) THEN
        cstate83 := 8; y1 := TRUE; t0_start := FALSE;t1_start := TRUE; t1_up := FALSE;
    ELSIF ((x1 = FALSE) AND  (t0.Q = FALSE) AND  ( TRUE )) THEN
        cstate83 := 1; y1 := FALSE; t0_start := FALSE;t1_start := FALSE;
    END_IF;
12:
    IF ((x1 = TRUE) AND  (t0.Q = TRUE) AND  ( TRUE )) THEN
        cstate83 := 9; y1 := FALSE; t0_start := TRUE; t0_up := FALSE;t1_start := FALSE;
    ELSIF ((x1 = FALSE) AND  ( TRUE ) AND  (t1.Q = FALSE)) THEN
        cstate83 := 16; y1 := FALSE; t0_start := FALSE;t1_start := FALSE;
    ELSIF ((x1 = TRUE) AND  (t0.Q = FALSE) AND  ( TRUE )) THEN
        cstate83 := 3; y1 := FALSE; t0_start := TRUE; t0_up := FALSE;t1_start := FALSE;
    ELSIF ((x1 = FALSE) AND  ( TRUE ) AND  (t1.Q = TRUE)) THEN
        cstate83 := 4; y1 := FALSE; t0_start := FALSE;t1_start := FALSE;
    END_IF;
13:
    IF ((x1 = TRUE) AND  (t0.Q = FALSE) AND  ( TRUE )) THEN
        cstate83 := 3; y1 := FALSE; t0_start := TRUE; t0_up := FALSE;t1_start := FALSE;
    ELSIF ((x1 = TRUE) AND  (t0.Q = TRUE) AND  ( TRUE )) THEN
        cstate83 := 9; y1 := FALSE; t0_start := TRUE; t0_up := FALSE;t1_start := FALSE;
    ELSIF ((x1 = FALSE) AND  ( TRUE ) AND  (t1.Q = TRUE)) THEN
        cstate83 := 4; y1 := FALSE; t0_start := FALSE;t1_start := FALSE;
    ELSIF ((x1 = FALSE) AND  ( TRUE ) AND  (t1.Q = FALSE)) THEN
        cstate83 := 16; y1 := FALSE; t0_start := FALSE;t1_start := FALSE;
    END_IF;
14:
    IF ((x1 = TRUE) AND  (t0.Q = FALSE) AND  (t1.Q = TRUE)) THEN
        cstate83 := 3; y1 := FALSE; t0_start := TRUE; t0_up := FALSE;t1_start := FALSE;
    ELSIF ((x1 = FALSE) AND  ( TRUE ) AND  (t1.Q = TRUE)) THEN
        cstate83 := 12; y1 := FALSE; t0_start := FALSE;t1_start := FALSE;
    ELSIF ((x1 = TRUE) AND  ( TRUE ) AND  (t1.Q = FALSE)) THEN
        cstate83 := 1; y1 := FALSE; t0_start := FALSE;t1_start := FALSE;
    ELSIF ((x1 = FALSE) AND  ( TRUE ) AND  (t1.Q = FALSE)) THEN
        cstate83 := 15; y1 := TRUE; t0_start := FALSE;t1_start := FALSE;
    ELSIF ((x1 = TRUE) AND  (t0.Q = TRUE) AND  (t1.Q = TRUE)) THEN
        cstate83 := 9; y1 := FALSE; t0_start := TRUE; t0_up := FALSE;t1_start := FALSE;
    END_IF;
15:
    IF ((x1 = TRUE) AND  (t0.Q = TRUE) AND  (t1.Q = TRUE)) THEN
        cstate83 := 9; y1 := FALSE; t0_start := TRUE; t0_up := FALSE;t1_start := FALSE;
    ELSIF ((x1 = FALSE) AND  ( TRUE ) AND  (t1.Q = TRUE)) THEN
        cstate83 := 12; y1 := FALSE; t0_start := FALSE;t1_start := FALSE;
    ELSIF ((x1 = TRUE) AND  (t0.Q = FALSE) AND  (t1.Q = TRUE)) THEN
        cstate83 := 3; y1 := FALSE; t0_start := TRUE; t0_up := FALSE;t1_start := FALSE;
    ELSIF ((x1 = TRUE) AND  ( TRUE ) AND  (t1.Q = FALSE)) THEN
        cstate83 := 1; y1 := FALSE; t0_start := FALSE;t1_start := FALSE;
    ELSIF ((x1 = FALSE) AND  ( TRUE ) AND  (t1.Q = FALSE)) THEN
        cstate83 := 15; y1 := TRUE; t0_start := FALSE;t1_start := FALSE;
    END_IF;
16:
    IF ((x1 = TRUE) AND  (t0.Q = TRUE) AND  ( TRUE )) THEN
        cstate83 := 9; y1 := FALSE; t0_start := TRUE; t0_up := FALSE;t1_start := FALSE;
    ELSIF ((x1 = FALSE) AND  ( TRUE ) AND  (t1.Q = TRUE)) THEN
        cstate83 := 4; y1 := FALSE; t0_start := FALSE;t1_start := FALSE;
    ELSIF ((x1 = FALSE) AND  ( TRUE ) AND  (t1.Q = FALSE)) THEN
        cstate83 := 16; y1 := FALSE; t0_start := FALSE;t1_start := FALSE;
    ELSIF ((x1 = TRUE) AND  (t0.Q = FALSE) AND  ( TRUE )) THEN
        cstate83 := 3; y1 := FALSE; t0_start := TRUE; t0_up := FALSE;t1_start := FALSE;
    END_IF;
17:
    IF ((x1 = FALSE) AND  ( TRUE ) AND  (t1.Q = FALSE)) THEN
        cstate83 := 8; y1 := TRUE; t0_start := FALSE;t1_start := TRUE; t1_up := FALSE;
    ELSIF ((x1 = TRUE) AND  (t0.Q = FALSE) AND  ( TRUE )) THEN
        cstate83 := 6; y1 := FALSE; t0_start := FALSE;t1_start := FALSE;
    ELSIF ((x1 = FALSE) AND  ( TRUE ) AND  (t1.Q = TRUE)) THEN
        cstate83 := 14; y1 := TRUE; t0_start := FALSE;t1_start := TRUE; t1_up := FALSE;
    ELSIF ((x1 = TRUE) AND  (t0.Q = TRUE) AND  ( TRUE )) THEN
        cstate83 := 7; y1 := FALSE; t0_start := FALSE;t1_start := FALSE;
    END_IF;
0:
    IF ((x1 = TRUE) AND  (t0.Q = FALSE) AND  ( TRUE )) THEN
        cstate83 := 17; y1 := FALSE; t0_start := FALSE;t1_start := FALSE;
    ELSIF ((x1 = FALSE) AND  ( TRUE ) AND  (t1.Q = FALSE)) THEN
        cstate83 := 2; y1 := FALSE; t0_start := FALSE;t1_start := FALSE;
    ELSIF ((x1 = FALSE) AND  ( TRUE ) AND  (t1.Q = TRUE)) THEN
        cstate83 := 13; y1 := FALSE; t0_start := FALSE;t1_start := FALSE;
    ELSIF ((x1 = TRUE) AND  (t0.Q = TRUE) AND  ( TRUE )) THEN
        cstate83 := 5; y1 := FALSE; t0_start := FALSE;t1_start := FALSE;
    END_IF;
1:
    IF (( TRUE )) THEN
        cstate83 := 1; y1 := FALSE; t0_start := FALSE;t1_start := FALSE;
    END_IF;
2:
    IF ((x1 = TRUE) AND  (t0.Q = FALSE) AND  ( TRUE )) THEN
        cstate83 := 3; y1 := FALSE; t0_start := TRUE; t0_up := FALSE;t1_start := FALSE;
    ELSIF ((x1 = FALSE) AND  ( TRUE ) AND  (t1.Q = FALSE)) THEN
        cstate83 := 16; y1 := FALSE; t0_start := FALSE;t1_start := FALSE;
    ELSIF ((x1 = TRUE) AND  (t0.Q = TRUE) AND  ( TRUE )) THEN
        cstate83 := 9; y1 := FALSE; t0_start := TRUE; t0_up := FALSE;t1_start := FALSE;
    ELSIF ((x1 = FALSE) AND  ( TRUE ) AND  (t1.Q = TRUE)) THEN
        cstate83 := 4; y1 := FALSE; t0_start := FALSE;t1_start := FALSE;
    END_IF;
3:
    IF ((x1 = FALSE) AND  (t0.Q = FALSE) AND  ( TRUE )) THEN
        cstate83 := 1; y1 := FALSE; t0_start := FALSE;t1_start := FALSE;
    ELSIF ((x1 = TRUE) AND  (t0.Q = FALSE) AND  ( TRUE )) THEN
        cstate83 := 11; y1 := FALSE; t0_start := FALSE;t1_start := FALSE;
    ELSIF ((x1 = FALSE) AND  (t0.Q = TRUE) AND  (t1.Q = TRUE)) THEN
        cstate83 := 14; y1 := TRUE; t0_start := FALSE;t1_start := TRUE; t1_up := FALSE;
    ELSIF ((x1 = FALSE) AND  (t0.Q = TRUE) AND  (t1.Q = FALSE)) THEN
        cstate83 := 8; y1 := TRUE; t0_start := FALSE;t1_start := TRUE; t1_up := FALSE;
    ELSIF ((x1 = TRUE) AND  (t0.Q = TRUE) AND  ( TRUE )) THEN
        cstate83 := 10; y1 := FALSE; t0_start := FALSE;t1_start := FALSE;
    END_IF;
4:
    IF ((x1 = FALSE) AND  ( TRUE ) AND  (t1.Q = TRUE)) THEN
        cstate83 := 4; y1 := FALSE; t0_start := FALSE;t1_start := FALSE;
    ELSIF ((x1 = TRUE) AND  (t0.Q = TRUE) AND  ( TRUE )) THEN
        cstate83 := 9; y1 := FALSE; t0_start := TRUE; t0_up := FALSE;t1_start := FALSE;
    ELSIF ((x1 = FALSE) AND  ( TRUE ) AND  (t1.Q = FALSE)) THEN
        cstate83 := 16; y1 := FALSE; t0_start := FALSE;t1_start := FALSE;
    ELSIF ((x1 = TRUE) AND  (t0.Q = FALSE) AND  ( TRUE )) THEN
        cstate83 := 3; y1 := FALSE; t0_start := TRUE; t0_up := FALSE;t1_start := FALSE;
    END_IF;
5:
    IF ((x1 = TRUE) AND  (t0.Q = FALSE) AND  ( TRUE )) THEN
        cstate83 := 6; y1 := FALSE; t0_start := FALSE;t1_start := FALSE;
    ELSIF ((x1 = FALSE) AND  ( TRUE ) AND  (t1.Q = TRUE)) THEN
        cstate83 := 14; y1 := TRUE; t0_start := FALSE;t1_start := TRUE; t1_up := FALSE;
    ELSIF ((x1 = FALSE) AND  ( TRUE ) AND  (t1.Q = FALSE)) THEN
        cstate83 := 8; y1 := TRUE; t0_start := FALSE;t1_start := TRUE; t1_up := FALSE;
    ELSIF ((x1 = TRUE) AND  (t0.Q = TRUE) AND  ( TRUE )) THEN
        cstate83 := 7; y1 := TRUE; t0_start := FALSE;t1_start := FALSE;
    END_IF;
6:
    IF ((x1 = TRUE) AND  (t0.Q = TRUE) AND  ( TRUE )) THEN
        cstate83 := 7; y1 := FALSE; t0_start := FALSE;t1_start := FALSE;
    ELSIF ((x1 = TRUE) AND  (t0.Q = FALSE) AND  ( TRUE )) THEN
        cstate83 := 6; y1 := FALSE; t0_start := FALSE;t1_start := FALSE;
    ELSIF ((x1 = FALSE) AND  ( TRUE ) AND  (t1.Q = TRUE)) THEN
        cstate83 := 14; y1 := TRUE; t0_start := FALSE;t1_start := TRUE; t1_up := FALSE;
    ELSIF ((x1 = FALSE) AND  ( TRUE ) AND  (t1.Q = FALSE)) THEN
        cstate83 := 8; y1 := TRUE; t0_start := FALSE;t1_start := TRUE; t1_up := FALSE;
    END_IF;
7:
    IF ((x1 = FALSE) AND  ( TRUE ) AND  (t1.Q = FALSE)) THEN
        cstate83 := 8; y1 := TRUE; t0_start := FALSE;t1_start := TRUE; t1_up := FALSE;
    ELSIF ((x1 = FALSE) AND  ( TRUE ) AND  (t1.Q = TRUE)) THEN
        cstate83 := 14; y1 := TRUE; t0_start := FALSE;t1_start := TRUE; t1_up := FALSE;
    ELSIF ((x1 = TRUE) AND  (t0.Q = FALSE) AND  ( TRUE )) THEN
        cstate83 := 6; y1 := FALSE; t0_start := FALSE;t1_start := FALSE;
    ELSIF ((x1 = TRUE) AND  (t0.Q = TRUE) AND  ( TRUE )) THEN
        cstate83 := 7; y1 := TRUE; t0_start := FALSE;t1_start := FALSE;
    END_IF;
8:
    IF ((x1 = TRUE) AND  (t0.Q = TRUE) AND  (t1.Q = TRUE)) THEN
        cstate83 := 9; y1 := FALSE; t0_start := TRUE; t0_up := FALSE;t1_start := FALSE;
    ELSIF ((x1 = FALSE) AND  ( TRUE ) AND  (t1.Q = TRUE)) THEN
        cstate83 := 12; y1 := FALSE; t0_start := FALSE;t1_start := FALSE;
    ELSIF ((x1 = TRUE) AND  ( TRUE ) AND  (t1.Q = FALSE)) THEN
        cstate83 := 1; y1 := FALSE; t0_start := FALSE;t1_start := FALSE;
    ELSIF ((x1 = FALSE) AND  ( TRUE ) AND  (t1.Q = FALSE)) THEN
        cstate83 := 15; y1 := TRUE; t0_start := FALSE;t1_start := FALSE;
    ELSIF ((x1 = TRUE) AND  (t0.Q = FALSE) AND  (t1.Q = TRUE)) THEN
        cstate83 := 3; y1 := FALSE; t0_start := TRUE; t0_up := FALSE;t1_start := FALSE;
    END_IF;
9:
    IF ((x1 = TRUE) AND  (t0.Q = TRUE) AND  ( TRUE )) THEN
        cstate83 := 10; y1 := TRUE; t0_start := FALSE;t1_start := FALSE;
    ELSIF ((x1 = FALSE) AND  (t0.Q = FALSE) AND  ( TRUE )) THEN
        cstate83 := 1; y1 := FALSE; t0_start := FALSE;t1_start := FALSE;
    ELSIF ((x1 = FALSE) AND  (t0.Q = TRUE) AND  (t1.Q = TRUE)) THEN
        cstate83 := 14; y1 := TRUE; t0_start := FALSE;t1_start := TRUE; t1_up := FALSE;
    ELSIF ((x1 = TRUE) AND  (t0.Q = FALSE) AND  ( TRUE )) THEN
        cstate83 := 11; y1 := FALSE; t0_start := FALSE;t1_start := FALSE;
    ELSIF ((x1 = FALSE) AND  (t0.Q = TRUE) AND  (t1.Q = FALSE)) THEN
        cstate83 := 8; y1 := TRUE; t0_start := FALSE;t1_start := TRUE; t1_up := FALSE;
    END_IF;
10:
    IF ((x1 = TRUE) AND  (t0.Q = TRUE) AND  ( TRUE )) THEN
        cstate83 := 7; y1 := TRUE; t0_start := FALSE;t1_start := FALSE;
    ELSIF ((x1 = TRUE) AND  (t0.Q = FALSE) AND  ( TRUE )) THEN
        cstate83 := 6; y1 := FALSE; t0_start := FALSE;t1_start := FALSE;
    ELSIF ((x1 = FALSE) AND  ( TRUE ) AND  (t1.Q = TRUE)) THEN
        cstate83 := 14; y1 := TRUE; t0_start := FALSE;t1_start := TRUE; t1_up := FALSE;
    ELSIF ((x1 = FALSE) AND  ( TRUE ) AND  (t1.Q = FALSE)) THEN
        cstate83 := 8; y1 := TRUE; t0_start := FALSE;t1_start := TRUE; t1_up := FALSE;
    END_IF;
END_CASE;

(* Additional processing to handle clocks - in CODESYS, it only starts
    with rising edge and can not be placed inside IF statement *)
IF(t0_up = TRUE) THEN
    t0_reset := TRUE;
ELSIF(t0_start = TRUE AND t0_up = FALSE) THEN
    t0_up := TRUE;  t0_reset := FALSE;
END_IF
t0(IN:=t0_reset, PT:=T0_VALUE);
IF(t1_up = TRUE) THEN
    t1_reset := TRUE;
ELSIF(t1_start = TRUE AND t1_up = FALSE) THEN
    t1_up := TRUE;  t1_reset := FALSE;
END_IF
t1(IN:=t1_reset, PT:=T1_VALUE);

END_FUNCTION_BLOCK

(* ---- G4LTL_ST9.st ---- *)
FUNCTION_BLOCK FB_G4LTL

   (* Variable definition *)
   VAR_INPUT
      x0	: BOOL;
      x1	: BOOL;
   END_VAR
   VAR_OUTPUT
      y0	: BOOL;
   END_VAR
   VAR
   (* The total number of states equals to 1 *)
      cstate1	: LINT := 0;
   END_VAR

   (* Control logic *)
CASE cstate1 OF
0:
    IF ((x0 = FALSE) AND  ( TRUE )) OR ((x0 = TRUE) AND  (x1 = TRUE)) THEN
        cstate1 := 0; y0 := FALSE;
    ELSIF ((x0 = TRUE) AND  (x1 = FALSE)) THEN
        cstate1 := 0; y0 := TRUE;
    END_IF;
END_CASE;

END_FUNCTION_BLOCK

(* ---- IndustrialAuto1.st ---- *)
FUNCTION_BLOCK FB_G4LTL

   (* Variable definition *)
   VAR_INPUT
      x0	: BOOL;
      x1	: BOOL;
   END_VAR
   VAR_OUTPUT
      y0	: BOOL;
   END_VAR
   VAR
   (* The total number of states equals to 1 *)
      cstate57	: LINT := 0;
   END_VAR

   (* Control logic *)
CASE cstate57 OF
0:
    IF ((x0 = FALSE) AND  ( TRUE )) OR ((x0 = TRUE) AND  (x1 = TRUE)) THEN
        cstate57 := 0; y0 := FALSE;
    ELSIF ((x0 = TRUE) AND  (x1 = FALSE)) THEN
        cstate57 := 0; y0 := TRUE;
    END_IF;
END_CASE;

END_FUNCTION_BLOCK

(* ---- IndustrialAuto10.st ---- *)
FUNCTION_BLOCK FB_G4LTL

   (* Variable definition *)
   VAR_INPUT
      x0	: BOOL;
      x1	: BOOL;
      x2	: BOOL;
      x10	: BOOL;
   END_VAR
   VAR_OUTPUT
      y0	: BOOL;
      y1	: BOOL;
   END_VAR
   VAR
   (* The total number of states equals to 13 *)
      cstate59	: LINT := 0;
   END_VAR

   (* Control logic *)
CASE cstate59 OF
11:
    IF ((x0 = TRUE) AND  (x1 = FALSE) AND  (x2 = TRUE) AND  (x10 = FALSE)) THEN
        cstate59 := 9; y0 := TRUE; y1 := FALSE;
    ELSIF ((x0 = TRUE) AND  (x1 = TRUE) AND  (x2 = TRUE) AND  (x10 = FALSE)) THEN
        cstate59 := 10; y0 := FALSE; y1 := FALSE;
    ELSIF ((x0 = FALSE) AND  ( TRUE ) AND  ( TRUE ) AND  (x10 = TRUE)) THEN
        cstate59 := 4; y0 := FALSE; y1 := FALSE;
    ELSIF ((x0 = TRUE) AND  (x1 = FALSE) AND  (x2 = FALSE) AND  (x10 = FALSE)) THEN
        cstate59 := 5; y0 := TRUE; y1 := TRUE;
    ELSIF ((x0 = FALSE) AND  ( TRUE ) AND  (x2 = TRUE) AND  (x10 = FALSE)) THEN
        cstate59 := 6; y0 := FALSE; y1 := FALSE;
    ELSIF ((x0 = FALSE) AND  ( TRUE ) AND  (x2 = FALSE) AND  (x10 = FALSE)) THEN
        cstate59 := 11; y0 := FALSE; y1 := TRUE;
    ELSIF ((x0 = TRUE) AND  ( TRUE ) AND  ( TRUE ) AND  (x10 = TRUE)) THEN
        cstate59 := 7; y0 := FALSE; y1 := FALSE;
    ELSIF ((x0 = TRUE) AND  (x1 = TRUE) AND  (x2 = FALSE) AND  (x10 = FALSE)) THEN
        cstate59 := 12; y0 := FALSE; y1 := TRUE;
    END_IF;
12:
    IF ((x0 = FALSE) AND  ( TRUE ) AND  (x2 = FALSE) AND  (x10 = FALSE)) THEN
        cstate59 := 11; y0 := FALSE; y1 := TRUE;
    ELSIF ((x0 = FALSE) AND  ( TRUE ) AND  (x2 = TRUE) AND  (x10 = FALSE)) THEN
        cstate59 := 6; y0 := FALSE; y1 := FALSE;
    ELSIF ((x0 = FALSE) AND  ( TRUE ) AND  ( TRUE ) AND  (x10 = TRUE)) THEN
        cstate59 := 4; y0 := FALSE; y1 := FALSE;
    ELSIF ((x0 = TRUE) AND  ( TRUE ) AND  (x2 = FALSE) AND  (x10 = FALSE)) THEN
        cstate59 := 12; y0 := FALSE; y1 := TRUE;
    ELSIF ((x0 = TRUE) AND  ( TRUE ) AND  (x2 = TRUE) AND  (x10 = FALSE)) THEN
        cstate59 := 10; y0 := FALSE; y1 := FALSE;
    ELSIF ((x0 = TRUE) AND  ( TRUE ) AND  ( TRUE ) AND  (x10 = TRUE)) THEN
        cstate59 := 7; y0 := FALSE; y1 := FALSE;
    END_IF;
0:
    IF ((x0 = TRUE) AND  (x1 = FALSE) AND  ( TRUE ) AND  (x10 = FALSE)) OR ((x0 = TRUE) AND  (x1 = TRUE) AND  (x2 = TRUE) AND  (x10 = FALSE)) THEN
        cstate59 := 10; y0 := FALSE; y1 := FALSE;
    ELSIF ((x0 = TRUE) AND  (x1 = TRUE) AND  (x2 = FALSE) AND  (x10 = FALSE)) THEN
        cstate59 := 12; y0 := FALSE; y1 := TRUE;
    ELSIF ((x0 = FALSE) AND  (x1 = TRUE) AND  (x2 = FALSE) AND  (x10 = FALSE)) THEN
        cstate59 := 11; y0 := FALSE; y1 := TRUE;
    ELSIF ((x0 = TRUE) AND  ( TRUE ) AND  ( TRUE ) AND  (x10 = TRUE)) THEN
        cstate59 := 7; y0 := FALSE; y1 := FALSE;
    ELSIF ((x0 = FALSE) AND  ( TRUE ) AND  ( TRUE ) AND  (x10 = TRUE)) THEN
        cstate59 := 4; y0 := FALSE; y1 := FALSE;
    ELSIF ((x0 = FALSE) AND  (x1 = FALSE) AND  ( TRUE ) AND  (x10 = FALSE)) OR ((x0 = FALSE) AND  (x1 = TRUE) AND  (x2 = TRUE) AND  (x10 = FALSE)) THEN
        cstate59 := 6; y0 := FALSE; y1 := FALSE;
    END_IF;
1:
    IF ((x0 = TRUE) AND  (x1 = FALSE) AND  (x2 = TRUE) AND  (x10 = FALSE)) THEN
        cstate59 := 2; y0 := TRUE; y1 := FALSE;
    ELSIF ((x0 = TRUE) AND  (x1 = TRUE) AND  (x2 = FALSE) AND  (x10 = FALSE)) THEN
        cstate59 := 8; y0 := FALSE; y1 := TRUE;
    ELSIF ((x0 = TRUE) AND  (x1 = FALSE) AND  (x2 = FALSE) AND  (x10 = FALSE)) THEN
        cstate59 := 3; y0 := TRUE; y1 := TRUE;
    ELSIF ((x0 = FALSE) AND  ( TRUE ) AND  (x2 = FALSE) AND  (x10 = TRUE)) OR ((x0 = FALSE) AND  ( TRUE ) AND  (x2 = TRUE) AND  ( TRUE )) THEN
        cstate59 := 4; y0 := FALSE; y1 := FALSE;
    ELSIF ((x0 = FALSE) AND  ( TRUE ) AND  (x2 = FALSE) AND  (x10 = FALSE)) THEN
        cstate59 := 1; y0 := FALSE; y1 := TRUE;
    ELSIF ((x0 = TRUE) AND  (x1 = FALSE) AND  ( TRUE ) AND  (x10 = TRUE)) OR ((x0 = TRUE) AND  (x1 = TRUE) AND  (x2 = FALSE) AND  (x10 = TRUE)) OR ((x0 = TRUE) AND  (x1 = TRUE) AND  (x2 = TRUE) AND  ( TRUE )) THEN
        cstate59 := 7; y0 := FALSE; y1 := FALSE;
    END_IF;
2:
    IF ((x0 = TRUE) AND  (x1 = TRUE) AND  (x2 = FALSE) AND  (x10 = FALSE)) THEN
        cstate59 := 8; y0 := FALSE; y1 := TRUE;
    ELSIF ((x0 = FALSE) AND  (x1 = FALSE) AND  ( TRUE ) AND  ( TRUE )) OR ((x0 = FALSE) AND  (x1 = TRUE) AND  (x2 = FALSE) AND  (x10 = TRUE)) OR ((x0 = FALSE) AND  (x1 = TRUE) AND  (x2 = TRUE) AND  ( TRUE )) THEN
        cstate59 := 4; y0 := FALSE; y1 := FALSE;
    ELSIF ((x0 = FALSE) AND  (x1 = TRUE) AND  (x2 = FALSE) AND  (x10 = FALSE)) THEN
        cstate59 := 1; y0 := FALSE; y1 := TRUE;
    ELSIF ((x0 = TRUE) AND  (x1 = FALSE) AND  ( TRUE ) AND  (x10 = TRUE)) OR ((x0 = TRUE) AND  (x1 = TRUE) AND  (x2 = FALSE) AND  (x10 = TRUE)) OR ((x0 = TRUE) AND  (x1 = TRUE) AND  (x2 = TRUE) AND  ( TRUE )) THEN
        cstate59 := 7; y0 := FALSE; y1 := FALSE;
    ELSIF ((x0 = TRUE) AND  (x1 = FALSE) AND  ( TRUE ) AND  (x10 = FALSE)) THEN
        cstate59 := 2; y0 := TRUE; y1 := FALSE;
    END_IF;
3:
    IF ((x0 = FALSE) AND  ( TRUE ) AND  (x2 = FALSE) AND  (x10 = TRUE)) OR ((x0 = FALSE) AND  ( TRUE ) AND  (x2 = TRUE) AND  ( TRUE )) THEN
        cstate59 := 4; y0 := FALSE; y1 := FALSE;
    ELSIF ((x0 = TRUE) AND  (x1 = FALSE) AND  (x2 = FALSE) AND  (x10 = FALSE)) THEN
        cstate59 := 3; y0 := TRUE; y1 := TRUE;
    ELSIF ((x0 = TRUE) AND  (x1 = TRUE) AND  (x2 = FALSE) AND  (x10 = FALSE)) THEN
        cstate59 := 8; y0 := FALSE; y1 := TRUE;
    ELSIF ((x0 = FALSE) AND  ( TRUE ) AND  (x2 = FALSE) AND  (x10 = FALSE)) THEN
        cstate59 := 1; y0 := FALSE; y1 := TRUE;
    ELSIF ((x0 = TRUE) AND  (x1 = FALSE) AND  ( TRUE ) AND  (x10 = TRUE)) OR ((x0 = TRUE) AND  (x1 = TRUE) AND  (x2 = FALSE) AND  (x10 = TRUE)) OR ((x0 = TRUE) AND  (x1 = TRUE) AND  (x2 = TRUE) AND  ( TRUE )) THEN
        cstate59 := 7; y0 := FALSE; y1 := FALSE;
    ELSIF ((x0 = TRUE) AND  (x1 = FALSE) AND  (x2 = TRUE) AND  (x10 = FALSE)) THEN
        cstate59 := 2; y0 := TRUE; y1 := FALSE;
    END_IF;
4:
    IF ((x0 = FALSE) AND  (x1 = TRUE) AND  (x2 = FALSE) AND  (x10 = FALSE)) THEN
        cstate59 := 1; y0 := FALSE; y1 := TRUE;
    ELSIF ((x0 = TRUE) AND  (x1 = TRUE) AND  (x2 = FALSE) AND  (x10 = FALSE)) THEN
        cstate59 := 8; y0 := FALSE; y1 := TRUE;
    ELSIF ((x0 = FALSE) AND  (x1 = FALSE) AND  ( TRUE ) AND  ( TRUE )) OR ((x0 = FALSE) AND  (x1 = TRUE) AND  (x2 = FALSE) AND  (x10 = TRUE)) OR ((x0 = FALSE) AND  (x1 = TRUE) AND  (x2 = TRUE) AND  ( TRUE )) THEN
        cstate59 := 4; y0 := FALSE; y1 := FALSE;
    ELSIF ((x0 = TRUE) AND  (x1 = FALSE) AND  ( TRUE ) AND  (x10 = FALSE)) THEN
        cstate59 := 2; y0 := TRUE; y1 := FALSE;
    ELSIF ((x0 = TRUE) AND  (x1 = FALSE) AND  ( TRUE ) AND  (x10 = TRUE)) OR ((x0 = TRUE) AND  (x1 = TRUE) AND  (x2 = FALSE) AND  (x10 = TRUE)) OR ((x0 = TRUE) AND  (x1 = TRUE) AND  (x2 = TRUE) AND  ( TRUE )) THEN
        cstate59 := 7; y0 := FALSE; y1 := FALSE;
    END_IF;
5:
    IF ((x0 = FALSE) AND  ( TRUE ) AND  (x2 = TRUE) AND  (x10 = FALSE)) THEN
        cstate59 := 6; y0 := FALSE; y1 := FALSE;
    ELSIF ((x0 = TRUE) AND  ( TRUE ) AND  ( TRUE ) AND  (x10 = TRUE)) THEN
        cstate59 := 7; y0 := FALSE; y1 := FALSE;
    ELSIF ((x0 = FALSE) AND  ( TRUE ) AND  ( TRUE ) AND  (x10 = TRUE)) THEN
        cstate59 := 4; y0 := FALSE; y1 := FALSE;
    ELSIF ((x0 = TRUE) AND  (x1 = FALSE) AND  (x2 = FALSE) AND  (x10 = FALSE)) THEN
        cstate59 := 5; y0 := TRUE; y1 := TRUE;
    ELSIF ((x0 = TRUE) AND  (x1 = TRUE) AND  (x2 = TRUE) AND  (x10 = FALSE)) THEN
        cstate59 := 10; y0 := FALSE; y1 := FALSE;
    ELSIF ((x0 = FALSE) AND  ( TRUE ) AND  (x2 = FALSE) AND  (x10 = FALSE)) THEN
        cstate59 := 11; y0 := FALSE; y1 := TRUE;
    ELSIF ((x0 = TRUE) AND  (x1 = TRUE) AND  (x2 = FALSE) AND  (x10 = FALSE)) THEN
        cstate59 := 12; y0 := FALSE; y1 := TRUE;
    ELSIF ((x0 = TRUE) AND  (x1 = FALSE) AND  (x2 = TRUE) AND  (x10 = FALSE)) THEN
        cstate59 := 9; y0 := TRUE; y1 := FALSE;
    END_IF;
6:
    IF ((x0 = FALSE) AND  (x1 = TRUE) AND  (x2 = FALSE) AND  (x10 = FALSE)) THEN
        cstate59 := 11; y0 := FALSE; y1 := TRUE;
    ELSIF ((x0 = TRUE) AND  ( TRUE ) AND  ( TRUE ) AND  (x10 = TRUE)) THEN
        cstate59 := 7; y0 := FALSE; y1 := FALSE;
    ELSIF ((x0 = FALSE) AND  (x1 = FALSE) AND  ( TRUE ) AND  (x10 = FALSE)) OR ((x0 = FALSE) AND  (x1 = TRUE) AND  (x2 = TRUE) AND  (x10 = FALSE)) THEN
        cstate59 := 6; y0 := FALSE; y1 := FALSE;
    ELSIF ((x0 = TRUE) AND  (x1 = FALSE) AND  ( TRUE ) AND  (x10 = FALSE)) THEN
        cstate59 := 9; y0 := TRUE; y1 := FALSE;
    ELSIF ((x0 = TRUE) AND  (x1 = TRUE) AND  (x2 = TRUE) AND  (x10 = FALSE)) THEN
        cstate59 := 10; y0 := FALSE; y1 := FALSE;
    ELSIF ((x0 = FALSE) AND  ( TRUE ) AND  ( TRUE ) AND  (x10 = TRUE)) THEN
        cstate59 := 4; y0 := FALSE; y1 := FALSE;
    ELSIF ((x0 = TRUE) AND  (x1 = TRUE) AND  (x2 = FALSE) AND  (x10 = FALSE)) THEN
        cstate59 := 12; y0 := FALSE; y1 := TRUE;
    END_IF;
7:
    IF ((x0 = TRUE) AND  (x1 = TRUE) AND  (x2 = FALSE) AND  (x10 = FALSE)) THEN
        cstate59 := 8; y0 := FALSE; y1 := TRUE;
    ELSIF ((x0 = FALSE) AND  (x1 = TRUE) AND  (x2 = FALSE) AND  (x10 = FALSE)) THEN
        cstate59 := 1; y0 := FALSE; y1 := TRUE;
    ELSIF ((x0 = TRUE) AND  (x1 = FALSE) AND  ( TRUE ) AND  ( TRUE )) OR ((x0 = TRUE) AND  (x1 = TRUE) AND  (x2 = FALSE) AND  (x10 = TRUE)) OR ((x0 = TRUE) AND  (x1 = TRUE) AND  (x2 = TRUE) AND  ( TRUE )) THEN
        cstate59 := 7; y0 := FALSE; y1 := FALSE;
    ELSIF ((x0 = FALSE) AND  (x1 = FALSE) AND  ( TRUE ) AND  ( TRUE )) OR ((x0 = FALSE) AND  (x1 = TRUE) AND  (x2 = FALSE) AND  (x10 = TRUE)) OR ((x0 = FALSE) AND  (x1 = TRUE) AND  (x2 = TRUE) AND  ( TRUE )) THEN
        cstate59 := 4; y0 := FALSE; y1 := FALSE;
    END_IF;
8:
    IF ((x0 = FALSE) AND  ( TRUE ) AND  (x2 = FALSE) AND  (x10 = TRUE)) OR ((x0 = FALSE) AND  ( TRUE ) AND  (x2 = TRUE) AND  ( TRUE )) THEN
        cstate59 := 4; y0 := FALSE; y1 := FALSE;
    ELSIF ((x0 = TRUE) AND  ( TRUE ) AND  (x2 = FALSE) AND  (x10 = FALSE)) THEN
        cstate59 := 8; y0 := FALSE; y1 := TRUE;
    ELSIF ((x0 = FALSE) AND  ( TRUE ) AND  (x2 = FALSE) AND  (x10 = FALSE)) THEN
        cstate59 := 1; y0 := FALSE; y1 := TRUE;
    ELSIF ((x0 = TRUE) AND  ( TRUE ) AND  (x2 = FALSE) AND  (x10 = TRUE)) OR ((x0 = TRUE) AND  ( TRUE ) AND  (x2 = TRUE) AND  ( TRUE )) THEN
        cstate59 := 7; y0 := FALSE; y1 := FALSE;
    END_IF;
9:
    IF ((x0 = TRUE) AND  (x1 = TRUE) AND  (x2 = TRUE) AND  (x10 = FALSE)) THEN
        cstate59 := 10; y0 := FALSE; y1 := FALSE;
    ELSIF ((x0 = FALSE) AND  (x1 = FALSE) AND  ( TRUE ) AND  (x10 = FALSE)) OR ((x0 = FALSE) AND  (x1 = TRUE) AND  (x2 = TRUE) AND  (x10 = FALSE)) THEN
        cstate59 := 6; y0 := FALSE; y1 := FALSE;
    ELSIF ((x0 = TRUE) AND  ( TRUE ) AND  ( TRUE ) AND  (x10 = TRUE)) THEN
        cstate59 := 7; y0 := FALSE; y1 := FALSE;
    ELSIF ((x0 = FALSE) AND  (x1 = TRUE) AND  (x2 = FALSE) AND  (x10 = FALSE)) THEN
        cstate59 := 11; y0 := FALSE; y1 := TRUE;
    ELSIF ((x0 = FALSE) AND  ( TRUE ) AND  ( TRUE ) AND  (x10 = TRUE)) THEN
        cstate59 := 4; y0 := FALSE; y1 := FALSE;
    ELSIF ((x0 = TRUE) AND  (x1 = TRUE) AND  (x2 = FALSE) AND  (x10 = FALSE)) THEN
        cstate59 := 12; y0 := FALSE; y1 := TRUE;
    ELSIF ((x0 = TRUE) AND  (x1 = FALSE) AND  ( TRUE ) AND  (x10 = FALSE)) THEN
        cstate59 := 9; y0 := TRUE; y1 := FALSE;
    END_IF;
10:
    IF ((x0 = TRUE) AND  (x1 = TRUE) AND  (x2 = FALSE) AND  (x10 = FALSE)) THEN
        cstate59 := 12; y0 := FALSE; y1 := TRUE;
    ELSIF ((x0 = TRUE) AND  (x1 = FALSE) AND  ( TRUE ) AND  (x10 = FALSE)) OR ((x0 = TRUE) AND  (x1 = TRUE) AND  (x2 = TRUE) AND  (x10 = FALSE)) THEN
        cstate59 := 10; y0 := FALSE; y1 := FALSE;
    ELSIF ((x0 = FALSE) AND  ( TRUE ) AND  ( TRUE ) AND  (x10 = TRUE)) THEN
        cstate59 := 4; y0 := FALSE; y1 := FALSE;
    ELSIF ((x0 = FALSE) AND  (x1 = TRUE) AND  (x2 = FALSE) AND  (x10 = FALSE)) THEN
        cstate59 := 11; y0 := FALSE; y1 := TRUE;
    ELSIF ((x0 = FALSE) AND  (x1 = FALSE) AND  ( TRUE ) AND  (x10 = FALSE)) OR ((x0 = FALSE) AND  (x1 = TRUE) AND  (x2 = TRUE) AND  (x10 = FALSE)) THEN
        cstate59 := 6; y0 := FALSE; y1 := FALSE;
    ELSIF ((x0 = TRUE) AND  ( TRUE ) AND  ( TRUE ) AND  (x10 = TRUE)) THEN
        cstate59 := 7; y0 := FALSE; y1 := FALSE;
    END_IF;
END_CASE;

END_FUNCTION_BLOCK

(* ---- IndustrialAuto11.st ---- *)
FUNCTION_BLOCK FB_G4LTL

   (* Variable definition *)
   VAR_INPUT
      x1	: BOOL;
      x2	: BOOL;
   END_VAR
   VAR_OUTPUT
      y0	: BOOL;
      y1	: BOOL;
      y2	: BOOL;
   END_VAR
   VAR
   (* The total number of states equals to 6 *)
      cstate55	: LINT := 0;
   END_VAR

   (* Control logic *)
CASE cstate55 OF
0:
    IF ((x1 = FALSE) AND  (x2 = TRUE)) THEN
        cstate55 := 1; y0 := FALSE; y1 := FALSE; y2 := TRUE;
    ELSIF ((x1 = FALSE) AND  (x2 = FALSE)) THEN
        cstate55 := 2; y0 := FALSE; y1 := FALSE; y2 := TRUE;
    ELSIF ((x1 = TRUE) AND  (x2 = FALSE)) THEN
        cstate55 := 3; y0 := TRUE; y1 := TRUE; y2 := FALSE;
    ELSIF ((x1 = TRUE) AND  (x2 = TRUE)) THEN
        cstate55 := 5; y0 := FALSE; y1 := FALSE; y2 := FALSE;
    END_IF;
1:
    IF ((x1 = TRUE) AND  (x2 = FALSE)) THEN
        cstate55 := 3; y0 := TRUE; y1 := TRUE; y2 := FALSE;
    ELSIF ((x1 = TRUE) AND  (x2 = TRUE)) THEN
        cstate55 := 5; y0 := FALSE; y1 := FALSE; y2 := FALSE;
    ELSIF ((x1 = FALSE) AND  ( TRUE )) THEN
        cstate55 := 1; y0 := FALSE; y1 := FALSE; y2 := TRUE;
    END_IF;
2:
    IF ((x1 = TRUE) AND  (x2 = FALSE)) THEN
        cstate55 := 3; y0 := TRUE; y1 := TRUE; y2 := FALSE;
    ELSIF ((x1 = FALSE) AND  (x2 = TRUE)) THEN
        cstate55 := 1; y0 := FALSE; y1 := FALSE; y2 := TRUE;
    ELSIF ((x1 = TRUE) AND  (x2 = TRUE)) THEN
        cstate55 := 5; y0 := FALSE; y1 := FALSE; y2 := FALSE;
    ELSIF ((x1 = FALSE) AND  (x2 = FALSE)) THEN
        cstate55 := 2; y0 := FALSE; y1 := FALSE; y2 := TRUE;
    END_IF;
3:
    IF ((x1 = FALSE) AND  (x2 = TRUE)) THEN
        cstate55 := 4; y0 := FALSE; y1 := FALSE; y2 := TRUE;
    ELSIF (( TRUE ) AND  (x2 = FALSE)) THEN
        cstate55 := 3; y0 := TRUE; y1 := TRUE; y2 := FALSE;
    ELSIF ((x1 = TRUE) AND  (x2 = TRUE)) THEN
        cstate55 := 5; y0 := FALSE; y1 := FALSE; y2 := FALSE;
    END_IF;
4:
    IF ((x1 = TRUE) AND  (x2 = FALSE)) THEN
        cstate55 := 3; y0 := TRUE; y1 := TRUE; y2 := FALSE;
    ELSIF ((x1 = TRUE) AND  (x2 = TRUE)) THEN
        cstate55 := 5; y0 := FALSE; y1 := FALSE; y2 := FALSE;
    ELSIF ((x1 = FALSE) AND  ( TRUE )) THEN
        cstate55 := 4; y0 := FALSE; y1 := FALSE; y2 := TRUE;
    END_IF;
5:
    IF ((x1 = FALSE) AND  (x2 = FALSE)) THEN
        cstate55 := 5; y0 := FALSE; y1 := FALSE; y2 := FALSE;
    ELSIF ((x1 = TRUE) AND  (x2 = TRUE)) THEN
        cstate55 := 5; y0 := FALSE; y1 := FALSE; y2 := FALSE;
    ELSIF ((x1 = TRUE) AND  (x2 = FALSE)) THEN
        cstate55 := 3; y0 := TRUE; y1 := TRUE; y2 := FALSE;
    ELSIF ((x1 = FALSE) AND  (x2 = TRUE)) THEN
        cstate55 := 4; y0 := FALSE; y1 := FALSE; y2 := TRUE;
    END_IF;
END_CASE;

END_FUNCTION_BLOCK
